// TIA Portal V20 export
Screen "200PRBCompleteDisplay_1"  1276x673
  ScreenItem "sequenceControlFaceplate_Lite_1" at 392,557 size 641x64  Type=HmiFaceplateContainer
  ScreenItem "Title_ScreenOverview_X390_Y2" at 390,2 size 500x30  Type=HmiTextBox
  ScreenItem "Button_Back_1" at 2,2 size 90x60  Type=HmiButton
  ScreenItem "Line_Header_X0_Y64" at 0,64 size 1276x0  Type=HmiLine
  ScreenItem "Tec-Unit_LegendᆉY2" at 1183,2 size 90x60  Type=HmiButton
  ScreenItem "permanentareaborderrectangle" at 0,0 size 0x0  Type=HmiRectangle
  ScreenItem "Button_Back" at 2,4 size 90x60  Type=HmiButton
  ScreenItem "Title_ScreenOverview_X390_Y2_1" at 380,5 size 510x57  Type=HmiTextBox
  ScreenItem "面板容器_1" at 10,267 size 163x70  Type=HmiFaceplateContainer
  ScreenItem "面板容器_3" at 193,267 size 163x70  Type=HmiFaceplateContainer
  ScreenItem "面板容器_4" at 10,335 size 163x70  Type=HmiFaceplateContainer
  ScreenItem "面板容器_2" at 1090,4 size 88x58  Type=HmiFaceplateContainer
  ScreenItem "OPMode1_Blocked" at 1164,6 size 14x14  Type=HmiGraphicView
  ScreenItem "OPMode4_Foreground_Blocked_1" at 1018,4 size 88x58  Type=HmiGraphicView
